FUNCTION_BLOCK Recipe_2 (* Extracted Composite Function Block Type *)
  (* Standard: 61499-2 *)
  (* Version 10/13/2026, macie *)
  PACKAGE Main;
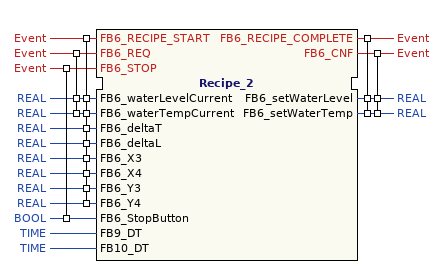
  EVENT_INPUT
    FB6_RECIPE_START WITH FB6_waterLevelCurrent, FB6_waterTempCurrent, FB6_deltaT, FB6_deltaL, FB6_X3, FB6_X4, FB6_Y3, FB6_Y4; (* Initialization Request *)
    FB6_REQ WITH FB6_waterLevelCurrent, FB6_waterTempCurrent; (* Normal Execution Request *)
    FB6_STOP WITH FB6_StopButton;
  END_EVENT
  EVENT_OUTPUT
    FB6_RECIPE_COMPLETE WITH FB6_setWaterLevel, FB6_setWaterTemp; (* Initialization Confirm *)
    FB6_CNF WITH FB6_setWaterLevel, FB6_setWaterTemp; (* Execution Confirmation *)
  END_EVENT
  VAR_INPUT
    FB6_waterLevelCurrent : REAL;
    FB6_waterTempCurrent : REAL; (* Input event qualifier *)
    FB6_deltaT : REAL;
    FB6_deltaL : REAL;
    FB6_X3 : REAL;
    FB6_X4 : REAL;
    FB6_Y3 : REAL;
    FB6_Y4 : REAL;
    FB6_StopButton : BOOL;
    FB9_DT : TIME; (* Delay Time *)
    FB10_DT : TIME; (* Delay Time *)
  END_VAR
  VAR_OUTPUT
    FB6_setWaterLevel : REAL; (* Output event qualifier *)
    FB6_setWaterTemp : REAL;
  END_VAR
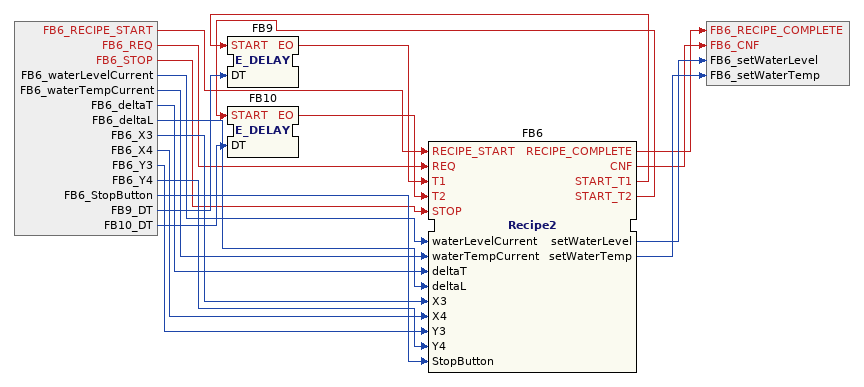
  FBS
    FB6 : Recipe2;
    FB9 : E_DELAY;
    FB10 : E_DELAY;
  END_FBS
  EVENT_CONNECTIONS
    FB10.EO TO FB6.T2;
    FB9.EO TO FB6.T1;
    FB6.START_T1 TO FB9.START;
    FB6.START_T2 TO FB10.START;
    FB6_RECIPE_START TO FB6.RECIPE_START;
    FB6_REQ TO FB6.REQ;
    FB6_STOP TO FB6.STOP;
    FB6.RECIPE_COMPLETE TO FB6_RECIPE_COMPLETE;
    FB6.CNF TO FB6_CNF;
  END_CONNECTIONS
  DATA_CONNECTIONS
    FB6_waterLevelCurrent TO FB6.waterLevelCurrent;
    FB6_waterTempCurrent TO FB6.waterTempCurrent;
    FB6_deltaT TO FB6.deltaT;
    FB6_deltaL TO FB6.deltaL;
    FB6_X3 TO FB6.X3;
    FB6_X4 TO FB6.X4;
    FB6_Y3 TO FB6.Y3;
    FB6_Y4 TO FB6.Y4;
    FB6_StopButton TO FB6.StopButton;
    FB6.setWaterLevel TO FB6_setWaterLevel;
    FB6.setWaterTemp TO FB6_setWaterTemp;
    FB9_DT TO FB9.DT;
    FB10_DT TO FB10.DT;
  END_CONNECTIONS
END_FUNCTION_BLOCK
